(* IEC 61131-3 sources: model-first-plc-agent-ai/results/T4-W-05, 2 files *)

(* ---- a1_code.st ---- *)
FUNCTION_BLOCK LevelControlRuntime
VAR_INPUT
    StartSignal : BOOL;
    StopSignal : BOOL;
    LevelValue : INT;
    ScaleValue : INT;
    h_span : REAL;
    h_sp : REAL;
    h_target : REAL;
    h_max : REAL;
    eps : REAL;
    t_h : TIME;
    Kp : REAL;
    Ti : REAL;
    Td : REAL;
    CycleSeconds : REAL;
END_VAR
VAR_OUTPUT
    FillCommand : INT;
    DischargeCommand : INT;
    fill_valve : BOOL;
    discharge_valve : BOOL;
END_VAR
VAR
    StartEdge : R_TRIG;
    HoldTimer : TON;

    start : BOOL;
    stop : BOOL;
    settled : BOOL;
    r : INT;

    x0 : BOOL := TRUE;
    x1 : BOOL := FALSE;

    h : REAL;
    ErrorValue : REAL;
    PreviousError : REAL := 0.0;
    IntegralTerm : REAL := 0.0;
    CandidateIntegral : REAL;
    DerivativeTerm : REAL;
    RawDemand : REAL;
    CandidateDemand : REAL;
    BoundedDemand : REAL;
    PidInitialized : BOOL := FALSE;
END_VAR

(* Region encoding: 0 = LOW, 1 = MID, 2 = HIGH. *)
StartEdge(CLK := StartSignal);
start := StartEdge.Q;
stop := StopSignal;

h := INT_TO_REAL(LevelValue) * h_span / INT_TO_REAL(ScaleValue);
ErrorValue := h_sp - h;

IF h < h_target THEN
    r := 0;
ELSIF h < h_max THEN
    r := 1;
ELSE
    r := 2;
END_IF;

(* The hold condition measures continuous time in tolerance in x1. *)
HoldTimer(
    IN := x1 AND NOT stop AND (ABS(ErrorValue) <= eps),
    PT := t_h
);
settled := HoldTimer.Q;

(* Evaluate transitions from the current situation only. *)
IF x0 THEN
    IF start AND NOT stop AND ((r = 0) OR (r = 1)) THEN
        x0 := FALSE;
        x1 := TRUE;
    END_IF;
ELSIF x1 THEN
    IF stop OR settled OR (r = 2) THEN
        x1 := FALSE;
        x0 := TRUE;
    END_IF;
ELSE
    x0 := TRUE;
    x1 := FALSE;
END_IF;

fill_valve := x1;
discharge_valve := x1;

FillCommand := 0;
DischargeCommand := 0;

IF fill_valve THEN
    (* Positional PID; demand is expressed as percent valve opening.
       Kp has units percent per level unit; Ti and Td are in seconds. *)
    IF NOT PidInitialized THEN
        PreviousError := ErrorValue;
        IntegralTerm := 0.0;
        PidInitialized := TRUE;
    END_IF;

    DerivativeTerm := 0.0;
    IF CycleSeconds > 0.0 THEN
        DerivativeTerm :=
            Kp * Td * (ErrorValue - PreviousError) / CycleSeconds;
    END_IF;

    RawDemand := Kp * ErrorValue + IntegralTerm + DerivativeTerm;

    (* Suspend integration whenever the current demand is clamped.
       Also reject an integral increment that would cause clamping. *)
    IF (RawDemand >= 0.0) AND (RawDemand <= 100.0)
       AND (Ti > 0.0) AND (CycleSeconds > 0.0) THEN
        CandidateIntegral :=
            IntegralTerm + Kp * ErrorValue * CycleSeconds / Ti;
        CandidateDemand :=
            Kp * ErrorValue + CandidateIntegral + DerivativeTerm;

        IF (CandidateDemand >= 0.0) AND (CandidateDemand <= 100.0) THEN
            IntegralTerm := CandidateIntegral;
            RawDemand := CandidateDemand;
        END_IF;
    END_IF;

    IF RawDemand < 0.0 THEN
        BoundedDemand := 0.0;
    ELSIF RawDemand > 100.0 THEN
        BoundedDemand := 100.0;
    ELSE
        BoundedDemand := RawDemand;
    END_IF;

    FillCommand :=
        REAL_TO_INT(BoundedDemand * INT_TO_REAL(ScaleValue) / 100.0);

    PreviousError := ErrorValue;
ELSE
    IntegralTerm := 0.0;
    PreviousError := ErrorValue;
    PidInitialized := FALSE;
    BoundedDemand := 0.0;
    settled := FALSE;
END_IF;

IF discharge_valve THEN
    DischargeCommand := REAL_TO_INT(0.4 * INT_TO_REAL(ScaleValue));
END_IF;

END_FUNCTION_BLOCK

PROGRAM Main
VAR
    StartCommand AT %IX100.0 : BOOL;
    StopCommand AT %IX100.1 : BOOL;
    LevelMeter AT %IW100 : INT;
    FillValve AT %QW100 : INT;
    DischargeValve AT %QW101 : INT;
END_VAR
VAR CONSTANT
    FULL_SCALE : INT := 1000;
END_VAR
VAR
    Controller : LevelControlRuntime;

    h_span : REAL := 10.0;
    h_sp : REAL;
    h_target : REAL;
    h_max : REAL;
    eps : REAL;
    t_h : TIME := T#10s;

    (* Initial tuning values; adjust for the simulated plant. *)
    Kp : REAL := 20.0;
    Ti : REAL := 5.0;
    Td : REAL := 0.0;

    (* Must match the configured periodic task interval. *)
    CycleSeconds : REAL := 0.02;
END_VAR

h_sp := 0.8 * h_span;
h_target := h_sp;
h_max := 0.9 * h_span;
eps := 0.02 * h_span;

Controller(
    StartSignal := StartCommand,
    StopSignal := StopCommand,
    LevelValue := LevelMeter,
    ScaleValue := FULL_SCALE,
    h_span := h_span,
    h_sp := h_sp,
    h_target := h_target,
    h_max := h_max,
    eps := eps,
    t_h := t_h,
    Kp := Kp,
    Ti := Ti,
    Td := Td,
    CycleSeconds := CycleSeconds
);

FillValve := Controller.FillCommand;
DischargeValve := Controller.DischargeCommand;

END_PROGRAM

CONFIGURATION Config0
    RESOURCE Res0 ON PLC
        TASK ControlTask(INTERVAL := T#20ms, PRIORITY := 0);
        PROGRAM MainInstance WITH ControlTask : Main;
    END_RESOURCE
END_CONFIGURATION

(* ---- a2_code.st ---- *)
FUNCTION_BLOCK FB_LevelControl
VAR_INPUT
    StartCommand : BOOL;
    StopCommand : BOOL;
    LevelMeter : INT;
    FullScaleValue : INT := 1000;
    h_span : REAL := 10.0;
    t_h : TIME := T#10s;
    Kp : REAL := 20.0;
    Ti : REAL := 5.0;
    Td : REAL := 0.0;
    CycleSeconds : REAL := 0.02;
END_VAR
VAR_OUTPUT
    FillValve : INT;
    DischargeValve : INT;
    fill_valve : BOOL;
    discharge_valve : BOOL;
END_VAR
VAR
    StartEdge : R_TRIG;
    HoldTimer : TON;
    start : BOOL;
    stop : BOOL;
    settled : BOOL;
    r : INT;
    SequenceState : INT := 0;
    x0 : BOOL := TRUE;
    x1 : BOOL := FALSE;
    WasRegulating : BOOL := FALSE;

    h : REAL;
    h_sp : REAL;
    h_target : REAL;
    h_max : REAL;
    eps : REAL;
    e : REAL;

    IntegralTerm : REAL := 0.0;
    PreviousError : REAL := 0.0;
    DerivativeTerm : REAL := 0.0;
    RawDemand : REAL := 0.0;
    BoundedDemand : REAL := 0.0;
    EffectiveCycle : REAL;
END_VAR
VAR CONSTANT
    R_LOW : INT := 0;
    R_MID : INT := 1;
    R_HIGH : INT := 2;
END_VAR

StartEdge(CLK := StartCommand);
start := StartEdge.Q;
stop := StopCommand;

EffectiveCycle := CycleSeconds;
IF EffectiveCycle <= 0.0 THEN
    EffectiveCycle := 0.02;
END_IF;

h_sp := 0.8 * h_span;
h_target := h_sp;
h_max := 0.9 * h_span;
eps := 0.02 * h_span;

IF FullScaleValue > 0 THEN
    h := INT_TO_REAL(LevelMeter) * h_span
         / INT_TO_REAL(FullScaleValue);
ELSE
    h := h_max;
END_IF;

e := h_sp - h;

IF h < h_target THEN
    r := R_LOW;
ELSIF h < h_max THEN
    r := R_MID;
ELSE
    r := R_HIGH;
END_IF;

(* Stop takes priority over starting or continuing regulation. *)
IF stop THEN
    SequenceState := 0;
ELSE
    CASE SequenceState OF
        0:
            IF start THEN
                SequenceState := 1;
            END_IF;
        1:
            SequenceState := 1;
    ELSE
        SequenceState := 0;
    END_CASE;
END_IF;

(* The hold interval is continuous and belongs to regulation only. *)
HoldTimer(
    IN := (SequenceState = 1) AND NOT stop AND (ABS(e) <= eps),
    PT := t_h
);
settled := HoldTimer.Q;

IF SequenceState = 1 THEN
    IF stop OR settled OR (r = R_HIGH) THEN
        SequenceState := 0;
    END_IF;
END_IF;

x0 := SequenceState = 0;
x1 := SequenceState = 1;
fill_valve := x1;
discharge_valve := x1;

FillValve := 0;
DischargeValve := 0;

IF x1 THEN
    (* Initialize the PID on entry without a derivative kick. *)
    IF NOT WasRegulating THEN
        IntegralTerm := 0.0;
        PreviousError := e;
    END_IF;

    DerivativeTerm := 0.0;
    IF Td > 0.0 THEN
        DerivativeTerm :=
            Kp * Td * (e - PreviousError) / EffectiveCycle;
    END_IF;

    IF Ti <= 0.0 THEN
        IntegralTerm := 0.0;
    END_IF;

    (* Demand is expressed in percent; error is expressed in volts. *)
    RawDemand := Kp * e + IntegralTerm + DerivativeTerm;

    IF RawDemand > 100.0 THEN
        BoundedDemand := 100.0;
    ELSIF RawDemand < 0.0 THEN
        BoundedDemand := 0.0;
    ELSE
        BoundedDemand := RawDemand;

        (* Suspend integration whenever the output is clamped. *)
        IF Ti > 0.0 THEN
            IntegralTerm :=
                IntegralTerm + Kp * e * EffectiveCycle / Ti;
        END_IF;
    END_IF;

    PreviousError := e;

    IF FullScaleValue > 0 THEN
        FillValve := REAL_TO_INT(
            BoundedDemand * INT_TO_REAL(FullScaleValue) / 100.0
        );
        DischargeValve := REAL_TO_INT(
            0.4 * INT_TO_REAL(FullScaleValue)
        );
    END_IF;
ELSE
    IntegralTerm := 0.0;
    PreviousError := e;
    DerivativeTerm := 0.0;
    RawDemand := 0.0;
    BoundedDemand := 0.0;

    (* Clear the owned hold condition immediately on leaving regulation. *)
    HoldTimer(IN := FALSE, PT := t_h);
    settled := FALSE;
END_IF;

WasRegulating := x1;

END_FUNCTION_BLOCK

PROGRAM Main
VAR
    StartCommand AT %IX100.0 : BOOL;
    StopCommand AT %IX100.1 : BOOL;
    LevelMeter AT %IW100 : INT;
    FillValve AT %QW100 : INT;
    DischargeValve AT %QW101 : INT;
END_VAR
VAR
    Controller : FB_LevelControl;
    Kp : REAL := 20.0;
    Ti : REAL := 5.0;
    Td : REAL := 0.0;
END_VAR
VAR CONSTANT
    FULL_SCALE : INT := 1000;
    h_span : REAL := 10.0;
    t_h : TIME := T#10s;
    CycleSeconds : REAL := 0.02;
END_VAR

Controller(
    StartCommand := StartCommand,
    StopCommand := StopCommand,
    LevelMeter := LevelMeter,
    FullScaleValue := FULL_SCALE,
    h_span := h_span,
    t_h := t_h,
    Kp := Kp,
    Ti := Ti,
    Td := Td,
    CycleSeconds := CycleSeconds
);

FillValve := Controller.FillValve;
DischargeValve := Controller.DischargeValve;

END_PROGRAM

CONFIGURATION Config0
    RESOURCE Res0 ON PLC
        TASK ControlTask(INTERVAL := T#20ms, PRIORITY := 0);
        PROGRAM MainInstance WITH ControlTask : Main;
    END_RESOURCE
END_CONFIGURATION
